Fanuc KAREL source: kd00053.KL

-- PROVISIONAL review KL for V940-1; original PC SHA256 c4a9e902fd613f6e287f53ca2cbcebd36cc07456c9f81bc289d2e81257200584
-- Incomplete behavior may be omitted. Consult companion uncertainty JSON. Do not deploy.
PROGRAM KD00053
%NOLOCKGROUP
VAR
  I : INTEGER
  J : INTEGER
  B : BOOLEAN
  R : REAL
  S : STRING[80]
BEGIN
  -- V9_ZERO_TABLE_METADATA_HINT layout=0001; no indexed target words; source/name/runtime held
  -- UNRESOLVED_PC offsets 5-19; opcodes 21,9D,52,23
  -- UNRESOLVED_PC offsets 24-28; opcodes 7F
END KD00053
